Yaskawa INFORM job: M_SPLIT.JBI

/JOB
//NAME M_SPLIT
//POS
///NPOS 0,0,0,0,0,0
//INST
///DATE 2026/10/26 01:19
///COMM Generated using RoboDK
///ATTR SC,RW,RJ
///GROUP1 RB1
NOP
CALL JOB:SPLITTE
CALL JOB:SPLITTE2
CALL JOB:SPLITTE3
CALL JOB:SPLITTE4
END
